(* IEC 61131-3 sources: volt/packages/volt-lsp-iec/test-corpus/pro2193/Device/Plc Logic/Application/09 Misc/Library Manager/L_IC1P_ComponentDirectory, 20 files *)

(* ---- L_IC1P_COMPONENTINFODATAINFO.dut ---- *)
TYPE L_IC1P_COMPONENTINFODATAINFO :
STRUCT
	INDEX : UINT;
	SUBINDEX : USINT;
	CONFIG : USINT;
	PSDATA : POINTER TO STRING;
END_STRUCT
END_TYPE

(* ---- L_IC1P_COMPONENTINFODATASOURCE.dut ---- *)
TYPE L_IC1P_COMPONENTINFODATASOURCE :
STRUCT
	SERIALNUMBER : L_IC1P_ComponentInfoDataInfo;
	MANUFACTURER : L_IC1P_ComponentInfoDataInfo;
	SOFTWAREREVISION : L_IC1P_ComponentInfoDataInfo;
	HARDWAREREVISION : L_IC1P_ComponentInfoDataInfo;
	DEVICECLASS : L_IC1P_ComponentInfoDataInfo;
	PRODUCTCODE : L_IC1P_ComponentInfoDataInfo;
END_STRUCT
END_TYPE

(* ---- L_IC1P_COMPONENTINFOID.dut ---- *)
TYPE L_IC1P_COMPONENTINFOID :
(
	SERIALNUMBER := 3,
	MANUFACTURER := 5,
	SOFTWAREREVISION := 9,
	HARDWAREREVISION := 10,
	DEVICECLASS := 11,
	PRODUCTCODE := 13
);
END_TYPE

(* ---- L_IC1P_ICOMPONENTDATAPROVIDER.itf ---- *)
INTERFACE L_IC1P_ICOMPONENTDATAPROVIDER
END_INTERFACE

METHOD GETADDRESS : POINTER TO L_IC1P_ComponentHardware
END_METHOD

METHOD SETAUTOMATICUPDATE : BOOL
VAR_INPUT
	XAUTOMATICDATAUPDATE : BOOL;
END_VAR
END_METHOD

METHOD SETDATAUPDATED : BOOL
VAR_INPUT
	XDATAUPDATED : BOOL;
END_VAR
END_METHOD

METHOD SETDEVICECLASS : BOOL
VAR_INPUT
	SDEVICECLASS : STRING;
END_VAR
END_METHOD

METHOD SETHARDWAREREVISION : BOOL
VAR_INPUT
	SHARDWAREREVISION : STRING;
END_VAR
END_METHOD

METHOD SETMANUFACTURER : BOOL
VAR_INPUT
	SMANUFACTURER : STRING;
END_VAR
END_METHOD

METHOD SETPRODUCTCODE : BOOL
VAR_INPUT
	SPRODUCTCODE : STRING;
END_VAR
END_METHOD

METHOD SETSERIALNUMBER : BOOL
VAR_INPUT
	SSERIALNUMBER : STRING;
END_VAR
END_METHOD

METHOD SETSOFTWAREREVISION : BOOL
VAR_INPUT
	SSOFTWAREREVISION : STRING;
END_VAR
END_METHOD

METHOD UPDATEDATAELEMENT : BOOL
VAR_INPUT
	INFOID : L_IC1P_ComponentInfoId;
	SDATA : STRING;
END_VAR
END_METHOD

(* ---- GETBOOLEANPROPERTY.pou ---- *)
FUNCTION GETBOOLEANPROPERTY : BOOL
VAR_INPUT
	STKEY : WSTRING;
END_VAR
END_FUNCTION

(* ---- GETCOMPANY.pou ---- *)
FUNCTION GETCOMPANY : WSTRING
END_FUNCTION

(* ---- GETNUMBERPROPERTY.pou ---- *)
FUNCTION GETNUMBERPROPERTY : DINT
VAR_INPUT
	STKEY : WSTRING;
END_VAR
END_FUNCTION

(* ---- GETTEXTPROPERTY.pou ---- *)
FUNCTION GETTEXTPROPERTY : WSTRING
VAR_INPUT
	STKEY : WSTRING;
END_VAR
END_FUNCTION

(* ---- GETTEXTPROPERTY2.pou ---- *)
FUNCTION GETTEXTPROPERTY2 : POINTER TO WSTRING
VAR_INPUT
	STKEY : WSTRING;
END_VAR
END_FUNCTION

(* ---- GETTITLE.pou ---- *)
FUNCTION GETTITLE : WSTRING
END_FUNCTION

(* ---- GETVERSION.pou ---- *)
FUNCTION GETVERSION : VERSION
END_FUNCTION

(* ---- GETVERSIONPROPERTY.pou ---- *)
FUNCTION GETVERSIONPROPERTY : VERSION
VAR_INPUT
	STKEY : WSTRING;
END_VAR
END_FUNCTION

(* ---- L_IC1P_GETAPPNAME.pou ---- *)
FUNCTION L_IC1P_GETAPPNAME : STRING
VAR_IN_OUT
	SINSTANCESTRFULL : STRING(255);
END_VAR
END_FUNCTION

(* ---- L_IC1P_GETDEVICENAME.pou ---- *)
FUNCTION L_IC1P_GETDEVICENAME : STRING
VAR_IN_OUT
	SINSTANCESTRFULL : STRING(255);
END_VAR
END_FUNCTION

(* ---- GLOBALTEXTLIST.pou ---- *)
FUNCTION_BLOCK GLOBALTEXTLIST
VAR
	M_TEXTLISTFILE : STRING(255);
	_STNAMESPACE : STRING;
END_VAR
END_FUNCTION_BLOCK

(* ---- L_IC1P_COMPONENTHARDWARE.pou ---- *)
FUNCTION_BLOCK L_IC1P_COMPONENTHARDWARE
VAR_INPUT
	SDEVICECLASS : STRING;
	SMANUFACTURER : STRING;
	SPRODUCTCODE : STRING;
	SSERIALNUMBER : STRING;
	SHARDWAREREVISION : STRING;
	SSOFTWAREREVISION : STRING;
	XAUTOMATICDATAUPDATE : BOOL;
	XDATAAVAILABLE : BOOL;
END_VAR
END_FUNCTION_BLOCK

METHOD GETADDRESS : POINTER TO L_IC1P_ComponentHardware
END_METHOD

METHOD SETAUTOMATICUPDATE : BOOL
VAR_INPUT
	XAUTOMATICDATAUPDATE : BOOL;
END_VAR
END_METHOD

METHOD SETDATAUPDATED : BOOL
VAR_INPUT
	XDATAUPDATED : BOOL;
END_VAR
END_METHOD

METHOD SETDEVICECLASS : BOOL
VAR_INPUT
	SDEVICECLASS : STRING;
END_VAR
END_METHOD

METHOD SETHARDWAREREVISION : BOOL
VAR_INPUT
	SHARDWAREREVISION : STRING;
END_VAR
END_METHOD

METHOD SETMANUFACTURER : BOOL
VAR_INPUT
	SMANUFACTURER : STRING;
END_VAR
END_METHOD

METHOD SETPRODUCTCODE : BOOL
VAR_INPUT
	SPRODUCTCODE : STRING;
END_VAR
END_METHOD

METHOD SETSERIALNUMBER : BOOL
VAR_INPUT
	SSERIALNUMBER : STRING;
END_VAR
END_METHOD

METHOD SETSOFTWAREREVISION : BOOL
VAR_INPUT
	SSOFTWAREREVISION : STRING;
END_VAR
END_METHOD

METHOD UPDATEDATAELEMENT : BOOL
VAR_INPUT
	INFOID : L_IC1P_ComponentInfoId;
	SDATA : STRING;
END_VAR
END_METHOD

(* ---- L_IC1P_DEVICECONTROLLER.pou ---- *)
FUNCTION_BLOCK L_IC1P_DEVICECONTROLLER
VAR
	REGISTERONCOMPONENTDIRECTORY : L_IC1P_RegisterOnComponentDirectory;
	XCMPDATAHANDLINGNOTFINISHED : BOOL := TRUE;
	READCONTROLLERCMPINFO : L_IC1P_ReadControllerComponentInfo;
	SCOMPNAME : STRING(80) := '';
	SINSTANCESTRFULL : STRING(255);
END_VAR
END_FUNCTION_BLOCK

METHOD CYCLICCALL : INT
END_METHOD

METHOD GETCOMPNAME : BOOL
END_METHOD

METHOD READCMPINFO : BOOL
END_METHOD

METHOD FB_EXIT : BOOL
VAR_INPUT
	BINCOPYCODE : BOOL;
END_VAR
END_METHOD

METHOD FB_INIT : BOOL
VAR_INPUT
	BINITRETAINS : BOOL;
	BINCOPYCODE : BOOL;
END_VAR
END_METHOD

(* ---- L_IC1P_READCONTROLLERCOMPONENTINFO.pou ---- *)
FUNCTION_BLOCK L_IC1P_READCONTROLLERCOMPONENTINFO
VAR_INPUT
	XEXECUTE : BOOL;
END_VAR
VAR_OUTPUT
	XDONE : BOOL;
	XERROR : BOOL;
	XBUSY : BOOL;
	EERRORID : WORD;
END_VAR
VAR_IN_OUT
	REGISTERONCOMPONENTDIRECTORY : L_IC1P_RegisterOnComponentDirectory;
END_VAR
VAR
	XEXECUTEOLD : BOOL;
	ISTATE : INT;
	XWAITFORPARAMETERREADDONE : BOOL;
	READPARAMETER : L_IPAP_ParameterRead;
	SREADDATA : STRING;
	SREADDATAINT : STRING;
	BYSDORETRYCOUNTER : BYTE;
	IREADCOMPONENTDATASTATE : INT;
	BYNROFBYTE : BYTE;
	SDO_READ_TIME_OUT : UDINT := 5000;
	MAX_SDO_RETRIES : BYTE := 3;
	C_INIT_READERRORSDO : WORD := 1;
END_VAR
END_FUNCTION_BLOCK

METHOD ACYCLICACTION
END_METHOD

METHOD GETCOMPONENTINFOINDEX : WORD
VAR_INPUT
	DATASELECTION : UDINT;
END_VAR
VAR_OUTPUT
	USISUB : USINT;
	XISSTRING : BOOL;
END_VAR
END_METHOD

METHOD READCMPINFO : BOOL
VAR_IN_OUT
	REGISTERONCOMPONENTDIRECTORY : L_IC1P_RegisterOnComponentDirectory;
END_VAR
END_METHOD

(* ---- L_IC1P_REGISTERONCOMPONENTDIRECTORY.pou ---- *)
FUNCTION_BLOCK L_IC1P_REGISTERONCOMPONENTDIRECTORY
VAR_OUTPUT
	ITFHWDATAPROVIDER : L_IC1P_IComponentDataProvider;
END_VAR
VAR_IN_OUT
	SINSTANCESTRFULL : STRING(255);
	SCOMPNAME : STRING(80);
END_VAR
VAR
	ITFCALLBACK : CmpEventMgr.ICmpEventCallback;
	HINTERFACERESETDONE : SysTypes.RTS_IEC_HANDLE := SysTypes.RTS_INVALID_HANDLE;
	HEVENTRESETDONE : SysTypes.RTS_IEC_HANDLE := SysTypes.RTS_INVALID_HANDLE;
	HINTERFACEDOWNLOADDONE : SysTypes.RTS_IEC_HANDLE := SysTypes.RTS_INVALID_HANDLE;
	HEVENTONLINEDOWNLOADDONE : SysTypes.RTS_IEC_HANDLE := SysTypes.RTS_INVALID_HANDLE;
	WCNTRESETDONE : WORD;
	WCNTDOWNLOADDONE : WORD;
	PTYPENAME : POINTER TO STRING;
	COMPONENTINFODATASOURCE : L_IC1P_ComponentInfoDataSource;
	XCOMPINFOSOURCEAVAILABLE : BOOL;
	COMPINFOSOURCEAVAILABLE : BOOL;
	COMPONENTINFOSUPPORTED : BOOL;
END_VAR
END_FUNCTION_BLOCK

METHOD FB_REINIT : BOOL
END_METHOD

METHOD FINDCOMPONENT : BOOL
END_METHOD

METHOD GETCOMPONENTINFOSOURCE
VAR_INPUT
	INFOID : L_IC1P_ComponentInfoId;
END_VAR
VAR_OUTPUT
	INDEX : UINT;
	SUBINDEX : USINT;
	CONFIG : USINT;
	PSDATA : POINTER TO STRING;
END_VAR
END_METHOD

METHOD SETAUTOMATICUPDATEAVAILABLE : BOOL
VAR_INPUT
	XAUTOMATICUPDATEAVAILABLE : BOOL;
END_VAR
END_METHOD

METHOD SETCOMPINFOSOURCEAVAILABLE : BOOL
VAR_INPUT
	XAVAILABLE : BOOL;
END_VAR
END_METHOD

METHOD SETCOMPONENTINFOSOURCE
VAR_INPUT
	INFOID : L_IC1P_ComponentInfoId;
	INDEX : UINT;
	SUBINDEX : USINT;
	CONFIG : USINT;
	PSDATA : POINTER TO STRING;
END_VAR
END_METHOD

METHOD FB_EXIT : BOOL
VAR_INPUT
	BINCOPYCODE : BOOL;
END_VAR
END_METHOD

METHOD FB_INIT : BOOL
VAR_INPUT
	BINITRETAINS : BOOL;
	BINCOPYCODE : BOOL;
END_VAR
END_METHOD

METHOD EVENTCALLBACK : UDINT
VAR_INPUT
	PEVENTPARAM : POINTER TO EventParam;
END_VAR
END_METHOD

METHOD REGISTEREVENT
VAR_INPUT
	XONLYCALLBACKFUNCTION : BOOL;
END_VAR
END_METHOD

METHOD UNREGISTEREVENT
VAR_INPUT
	XONLYCALLBACKFUNCTION : BOOL;
END_VAR
END_METHOD

(* ---- L_IC1P_SYMBOLCONFIG.pou ---- *)
FUNCTION_BLOCK L_IC1P_SYMBOLCONFIG
VAR
	_VARACCESSIBASE : IecVarAccessLibrary.IBase;
	_PPIVARACCESS3 : POINTER TO IecVarAccessLibrary.IIecVarAccess3;
	_VARACCESS3 : IecVarAccessLibrary.IIecVarAccess3;
	_PPIVARACCESS4 : POINTER TO IecVarAccessLibrary.IIecVarAccess4;
	_VARACCESS4 : IecVarAccessLibrary.IIecVarAccess4;
	_PPIVARACCESS5 : POINTER TO IecVarAccessLibrary.IIecVarAccess5;
	_VARACCESS5 : IecVarAccessLibrary.IIecVarAccess5;
	_PPIVARACCESS7 : POINTER TO IecVarAccessLibrary.IIecVarAccess7;
	_VARACCESS7 : IecVarAccessLibrary.IIecVarAccess7;
	_SSYMBOL : STRING(255);
	_HNODE : IecVarAccessLibrary.ICollections.IBaseTreeNode;
	_VARINFO : VariableInformationStruct;
END_VAR
END_FUNCTION_BLOCK

METHOD GETADDRESS : POINTER TO BYTE
VAR_OUTPUT
	RESULT : SysTypes.RTS_IEC_RESULT;
END_VAR
END_METHOD

METHOD GETTYPENAME : POINTER TO STRING
END_METHOD

METHOD INIT : BOOL
VAR_IN_OUT
	RESULT : SysTypes.RTS_IEC_RESULT;
END_VAR
END_METHOD

METHOD REQUEST : BOOL
VAR_INPUT
	SSYMBOL : STRING(255);
END_VAR
END_METHOD
